(* PLC project TBEN_L5_PLC11.project, CODESYS CODESYS V3.5 SP21 Patch 1 *)
(* stored: creationDateTime 2026-11-07T15:35:08.8307014, modificationDateTime 2026-11-07T15:09:07.4034196 *)

// TRUE nếu STATUS RDREC/WRREC là "state conflict" (B5) hoặc "resource busy" (C3) -> master chưa xong, được retry
FUNCTION F_IolIsPnioBusy : BOOL
VAR_INPUT
    dwStatus : DWORD;          // ErrorCode, ErrorDecode, ErrorCode1, ErrorCode2 (byte cao -> thấp)
END_VAR
VAR
    bCode1 : BYTE;
END_VAR

            bCode1 := DWORD_TO_BYTE(SHR(dwStatus, 8));
F_IolIsPnioBusy := (bCode1 = 16#B5) OR (bCode1 = 16#C3);

          
END_FUNCTION
